(* PLC project g_vessel_empty_permissive_bomb, Anonymous Benchmark Suite 1.0 *)
(* stored: creationDateTime 2026-09-02T00:00:00 *)

PROGRAM g_vessel_empty_permissive_bomb
  VAR_INPUT
    feed_cmd : BOOL;
    discharge_cmd : BOOL;
    vessel_empty : BOOL;
    maint : BOOL;
  END_VAR
  VAR_OUTPUT
    feed_valve : BOOL;
    discharge_valve : BOOL;
  END_VAR

(* LD diagram, written out as Structured Text *)
feed_valve := NOT discharge_cmd AND vessel_empty AND feed_cmd OR feed_cmd AND maint;
discharge_valve := discharge_cmd AND NOT vessel_empty;
END_PROGRAM

CONFIGURATION Config0
  RESOURCE Res0 ON PLC
    TASK tcyclic(INTERVAL := T#10ms, PRIORITY := 0);
    PROGRAM inst0 WITH tcyclic : g_vessel_empty_permissive_bomb;
  END_RESOURCE
END_CONFIGURATION
